(* IEC 61131-3 sources: virtual-bottling-plant/plc/src/types, 2 files *)

(* ---- ST_MachineCmd.st ---- *)
(* One-scan PackML commands to one machine (from FB_LineSequencer). *)
TYPE
  ST_MachineCmd : STRUCT
    Start : BOOL;
    Stop : BOOL;
    Reset : BOOL;   (* Stopped → Idle, and Held → Unholding (unhold) *)
    Abort : BOOL;
    Clear : BOOL;
  END_STRUCT;
END_TYPE

(* ---- ST_Recipe.st ---- *)
(* Active recipe in the PLC (PLC-30). Written only by FB_RecipeHandshake. *)
TYPE
  ST_Recipe : STRUCT
    RecipeId : INT;
    RecipeVersion : INT;
    ProductCode : INT;      (* 1 = orange, 2 = apple *)
    BrixTarget : REAL;      (* °Bx *)
    BrixTol : REAL;         (* ± °Bx *)
    ConcRatio : REAL;       (* L concentrate per L of batch *)
    FillTargetG : REAL;     (* g per bottle *)
    LineSpeed : REAL;       (* bpm at the filler, the line constraint *)
    CapTorque : REAL;       (* Nm *)
  END_STRUCT;
END_TYPE
